// SIMATIC S7-200 SMART project (STEP 7-Micro/WIN SMART), CPU ST20

SYMBOL_TABLE 表格 1
Btn_set_Charge   V536.3
Calc_Temp_Real   VD700    // 计算中间暂存区 (DInt/Real)
Comm_State_Counter VB548    // 串口发送逻辑切换计数器
Comm_State_Counter1 VB549
HMI_IP_Apply     V536.2   // HMI 确认修改 IP 按钮
HMI_Start_Btn    V536.0   // HMI 手动开始按钮
HMI_Stop_Btn     V536.1   // HMI 手动停止按钮
Input_Current    VD504    // 实时输入电流 (A)
Input_Power      VD508    // 实时输入功率 (W)
Input_Voltage    VD500    // 实时输入电压 (V)
Output_Current   VD516    // 实时输出电流 (A)
Output_Voltage   VD512    // 实时输出电压 (V)
PLC_IP_Octet1    VB908    // PLC IP 地址第 1 段
PLC_IP_Octet2    VB909    // PLC IP 地址第 2 段
PLC_IP_Octet3    VB910    // PLC IP 地址第 3 段
PLC_IP_Octet4    VB911    // PLC IP 地址第 4 段
PN_In_Cmd        IB1160   // PN 接收自 1200: 远程启停指令
PN_In_SetI       ID1156   // PN 接收自 1200: 远程设定电流
PN_In_SetV       ID1152   // PN 接收自 1200: 远程设定电压
PN_Out_Curr      QD1156   // PN 发送给 1200: 输出电流
PN_Out_SetI      QD1164   // PN 发送给 1200: 当前设定电流
PN_Out_SetV      QD1160   // PN 发送给 1200: 当前设定电压
PN_Out_Status    QB1168   // PN 发送给 1200: 系统状态字节
PN_Out_Volt      QD1152   // PN 发送给 1200: 输出电压
Set_Current      VD532    // HMI 设定电流值 (默认 15.0)
Set_Voltage      VD528    // HMI 设定电压值 (默认 54.0)
Status_Bat_FB    V537.2   // 电池接入状态 (对应 Q0.1)
Status_Fault_FB  V537.1   // 系统故障状态 (对应 Q0.2)
Status_Run_FB    V537.0   // 充电运行状态 (对应 Q0.0)
Status_开关机标志     V537.3
Temp_T1          VD520    // 模块温度 T1 (℃)
Temp_T2          VD524    // 模块温度 T2 (℃)
发送数据             VB600    // 串口发送缓冲区起始 (长度 13)
启动接收并存入_VB550    VB550
END_SYMBOL_TABLE

SYMBOL_TABLE 系统符号
Always_On        SM0.0    // 始终接通
First_Scan_On    SM0.1    // 仅在第一个扫描周期时接通
P0_Config        SMB30    // 组态端口 0 通信：奇偶校验、每个字符的数据位数、波特率和协议
P0_Ctrl_Rcv      SMB87    // 接收消息控制
P0_End_Char      SMB89    // 消息结束字符
P0_Timeout       SMW92    // 字符间/消息定时器超时值，以毫秒为单位指定
P0_Max_Char      SMB94    // 要接收的最大字符数（1 到 255 字节）
END_SYMBOL_TABLE

ORGANIZATION_BLOCK MAIN:OB1
TITLE=
BEGIN
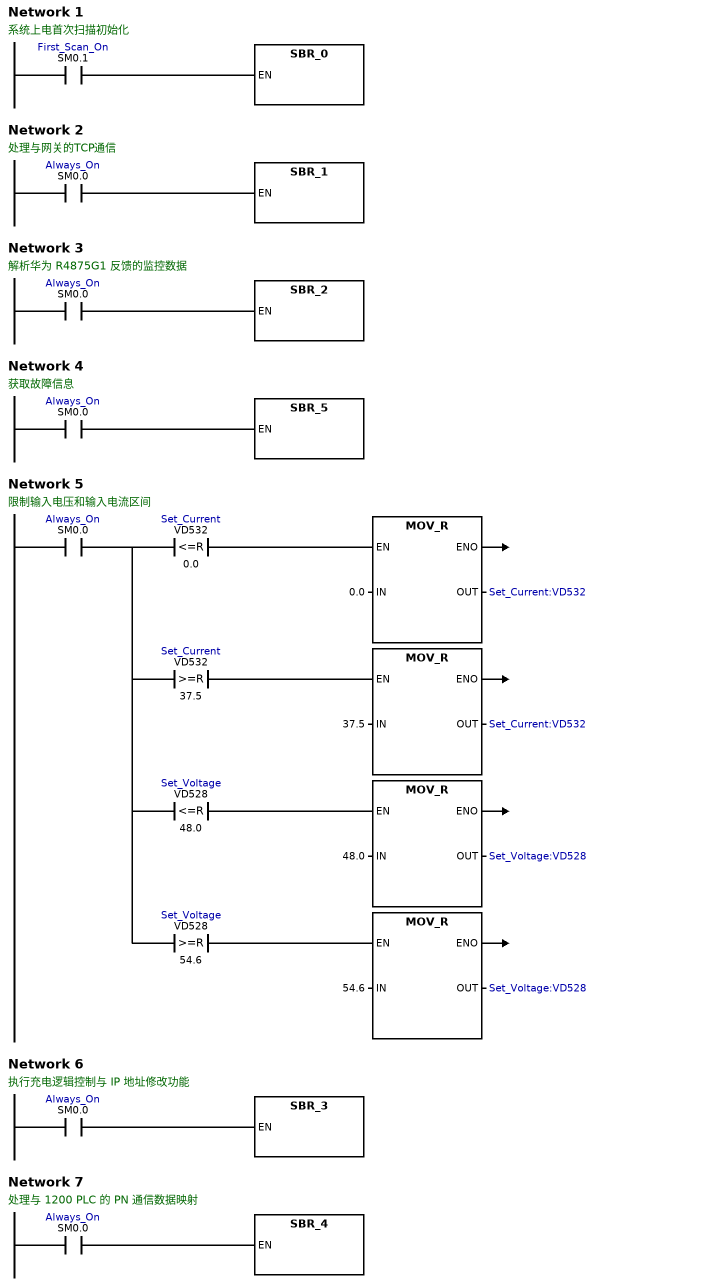
Network 1
//  系统上电首次扫描初始化
// 载入首次扫描标志位
// 调用初始化子程序
LD     First_Scan_On:SM0.1
CALL   SBR_0:SBR0
Network 2
//  处理与网关的TCP通信
// 始终接通
// 调用通信子程序
LD     Always_On:SM0.0
CALL   SBR_1:SBR1
Network 3
//  解析华为 R4875G1 反馈的监控数据
// 始终接通
// 调用解析子程序
LD     Always_On:SM0.0
CALL   SBR_2:SBR2
Network 4
// 获取故障信息
// 始终接通
// 调用获取故障程序
LD     Always_On:SM0.0
CALL   SBR_5:SBR5
Network 5
// 限制输入电压和输入电流区间
LD     Always_On:SM0.0
LPS
AR<=   Set_Current:VD532, 0.0
MOVR   0.0, Set_Current:VD532
LRD
AR>=   Set_Current:VD532, 37.5
MOVR   37.5, Set_Current:VD532
LRD
AR<=   Set_Voltage:VD528, 48.0
MOVR   48.0, Set_Voltage:VD528
LPP
AR>=   Set_Voltage:VD528, 54.6
MOVR   54.6, Set_Voltage:VD528
Network 6
//  执行充电逻辑控制与 IP 地址修改功能
// 始终接通
// 调用控制子程序
LD     Always_On:SM0.0
CALL   SBR_3:SBR3
Network 7
//  处理与 1200 PLC 的 PN 通信数据映射
// 始终接通
// 调用通信映射子程序
LD     Always_On:SM0.0
CALL   SBR_4:SBR4
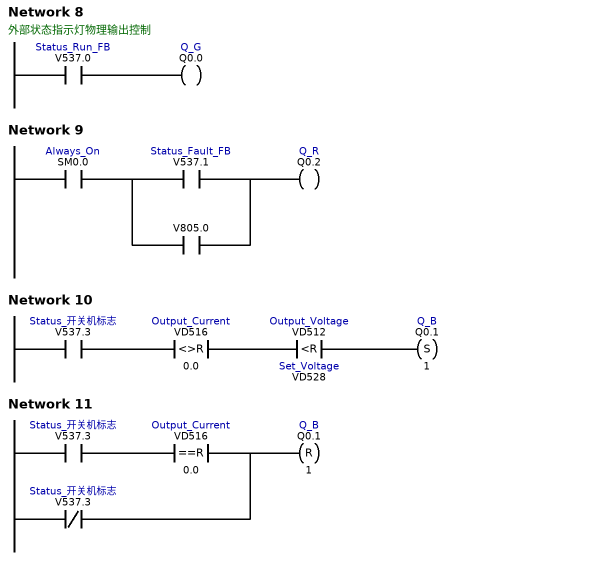
Network 8
//  外部状态指示灯物理输出控制
// 检查运行状态位
// 输出 Q0.0 绿灯: 充电运行
LD     Status_Run_FB:V537.0
=      Q_G:Q0.0
Network 9
// 检查故障状态位
// 输出 Q0.2 红灯: 系统故障
LD     Always_On:SM0.0
LD     Status_Fault_FB:V537.1
O      V805.0
ALD
=      Q_R:Q0.2
Network 10
// 检查电池接入位 (特殊标记：需用户自行完善)
// 输出 Q0.1 蓝灯: 电池接入
LD     Status_开关机标志:V537.3
AR<>   Output_Current:VD516, 0.0
AR<    Output_Voltage:VD512, Set_Voltage:VD528
S      Q_B:Q0.1, 1
Network 11
// 检查电池接入位 (特殊标记：需用户自行完善)
// 输出 Q0.1 蓝灯: 电池接入
LD     Status_开关机标志:V537.3
AR=    Output_Current:VD516, 0.0
ON     Status_开关机标志:V537.3
R      Q_B:Q0.1, 1
END_ORGANIZATION_BLOCK

SUBROUTINE_BLOCK SBR_0:SBR0
TITLE=初始化子程序
BEGIN
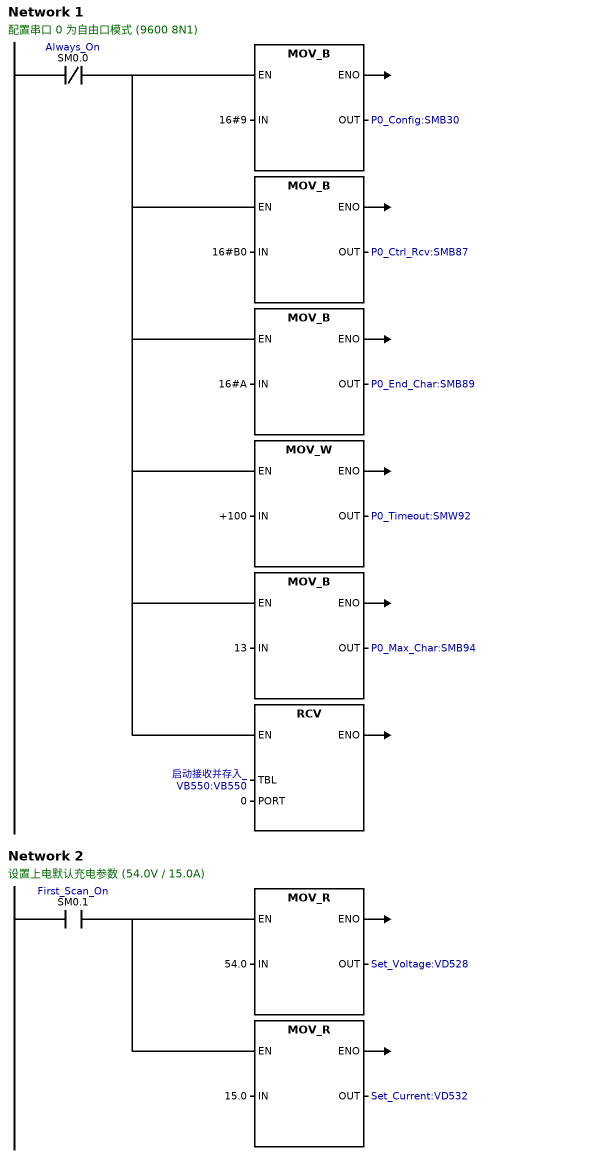
Network 1
//  配置串口 0 为自由口模式 (9600 8N1)
// 始终接通
// 端口 0: 9600, 8, N, 1, 自由口
// 设置接收控制: 允许接收, 超时结束
// 设置结束符 (0x0A)
// 设置接收超时 100ms
// 设置最大接收长度 13 字节
// 启动接收并存入 VB550
LDN    Always_On:SM0.0
MOVB   16#9, P0_Config:SMB30
MOVB   16#B0, P0_Ctrl_Rcv:SMB87
MOVB   16#A, P0_End_Char:SMB89
MOVW   +100, P0_Timeout:SMW92
MOVB   13, P0_Max_Char:SMB94
RCV    启动接收并存入_VB550:VB550, 0
Network 2
//  设置上电默认充电参数 (54.0V / 15.0A)
// 首次扫描
// 默认设定电压 54.0V
// 默认设定电流 15.0A
LD     First_Scan_On:SM0.1
MOVR   54.0, Set_Voltage:VD528
MOVR   15.0, Set_Current:VD532
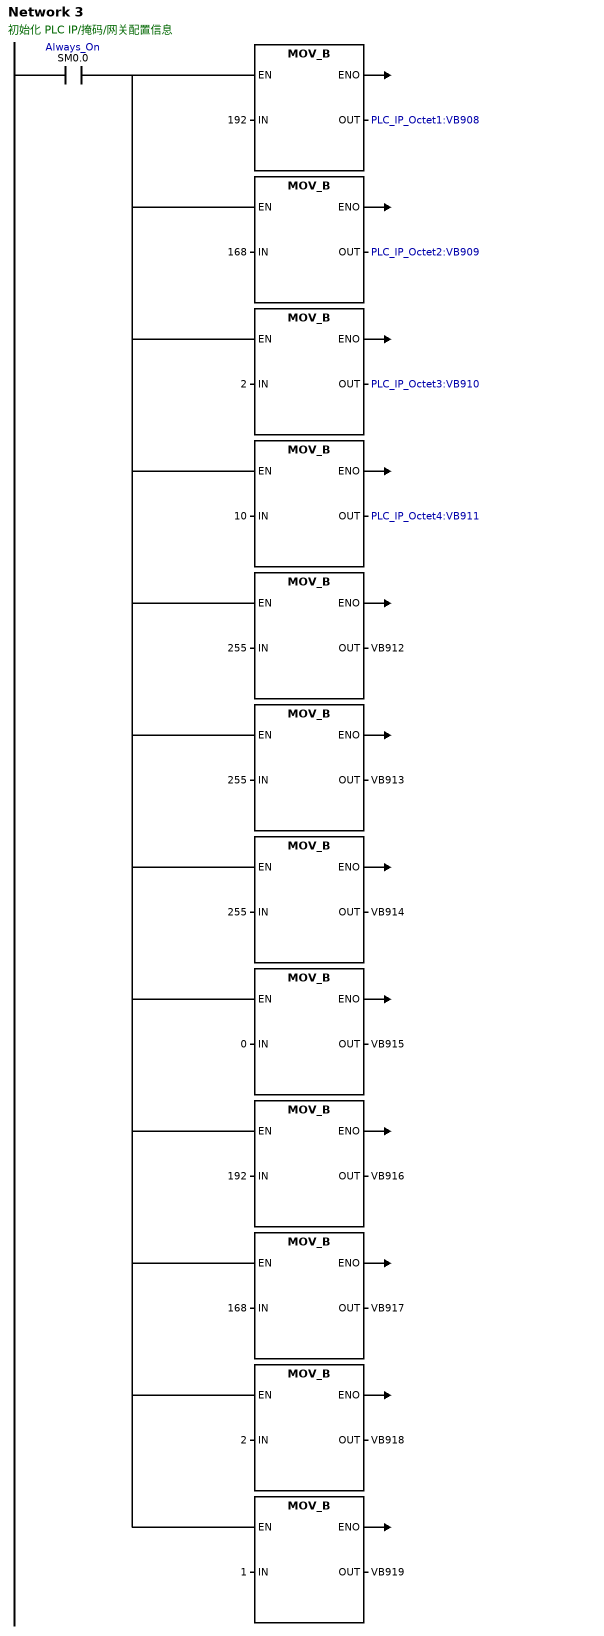
Network 3
//  初始化 PLC IP/掩码/网关配置信息
// 首次扫描
// IP 第一段
// IP 第二段
// IP 第三段
// IP 第四段
// 掩码第一段
// 掩码第二段
// 掩码第三段
// 掩码第四段
// 网关第一段
// 网关第二段
// 网关第三段
// 网关第四段
LD     Always_On:SM0.0
MOVB   192, PLC_IP_Octet1:VB908
MOVB   168, PLC_IP_Octet2:VB909
MOVB   2, PLC_IP_Octet3:VB910
MOVB   10, PLC_IP_Octet4:VB911
MOVB   255, VB912
MOVB   255, VB913
MOVB   255, VB914
MOVB   0, VB915
MOVB   192, VB916
MOVB   168, VB917
MOVB   2, VB918
MOVB   1, VB919
END_SUBROUTINE_BLOCK

SUBROUTINE_BLOCK SBR_1:SBR1
TITLE=TCP通信 - 华为协议
BEGIN
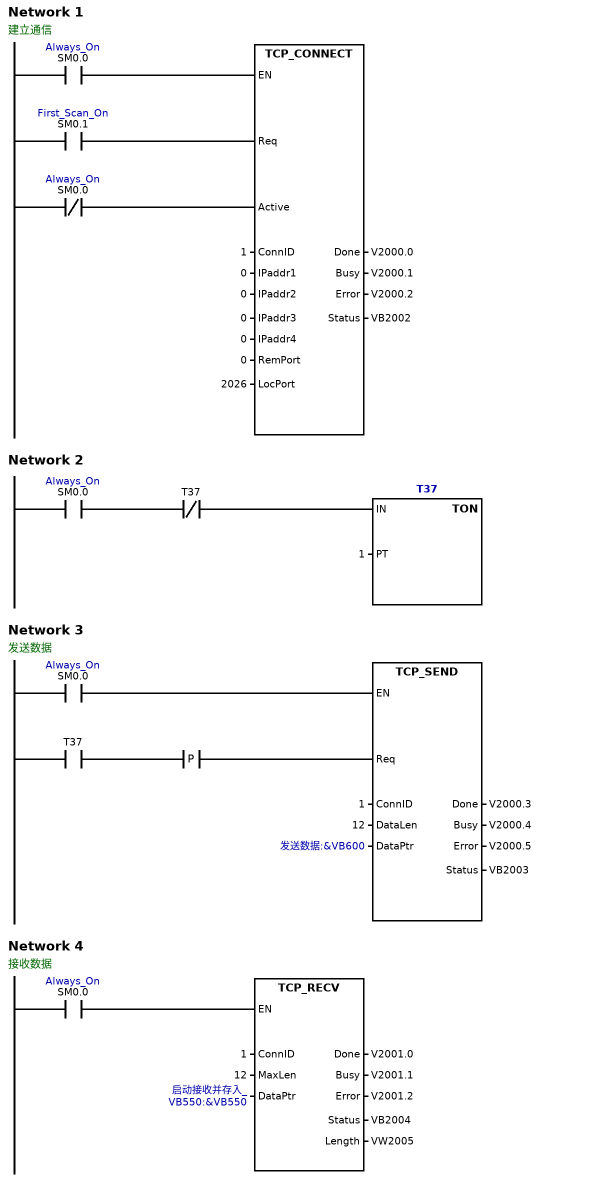
Network 1
// 建立通信
LD     Always_On:SM0.0
=      L60.0
LD     First_Scan_On:SM0.1
=      L63.7
LDN    Always_On:SM0.0
=      L63.6
LD     L60.0
CALL   TCP_CONNECT:SBR6, L63.7, L63.6, 1, 0, 0, 0, 0, 0, 2026, V2000.0, V2000.1, V2000.2, VB2002
Network 2
LD     Always_On:SM0.0
AN     T37
TON    T37, 1
Network 3
// 发送数据
LD     Always_On:SM0.0
=      L60.0
LD     T37
EU
=      L63.7
LD     L60.0
CALL   TCP_SEND:SBR7, L63.7, 1, 12, &发送数据:VB600, V2000.3, V2000.4, V2000.5, VB2003
Network 4
// 接收数据
LD     Always_On:SM0.0
CALL   TCP_RECV:SBR8, 1, 12, &启动接收并存入_VB550:VB550, V2001.0, V2001.1, V2001.2, VB2004, VW2005
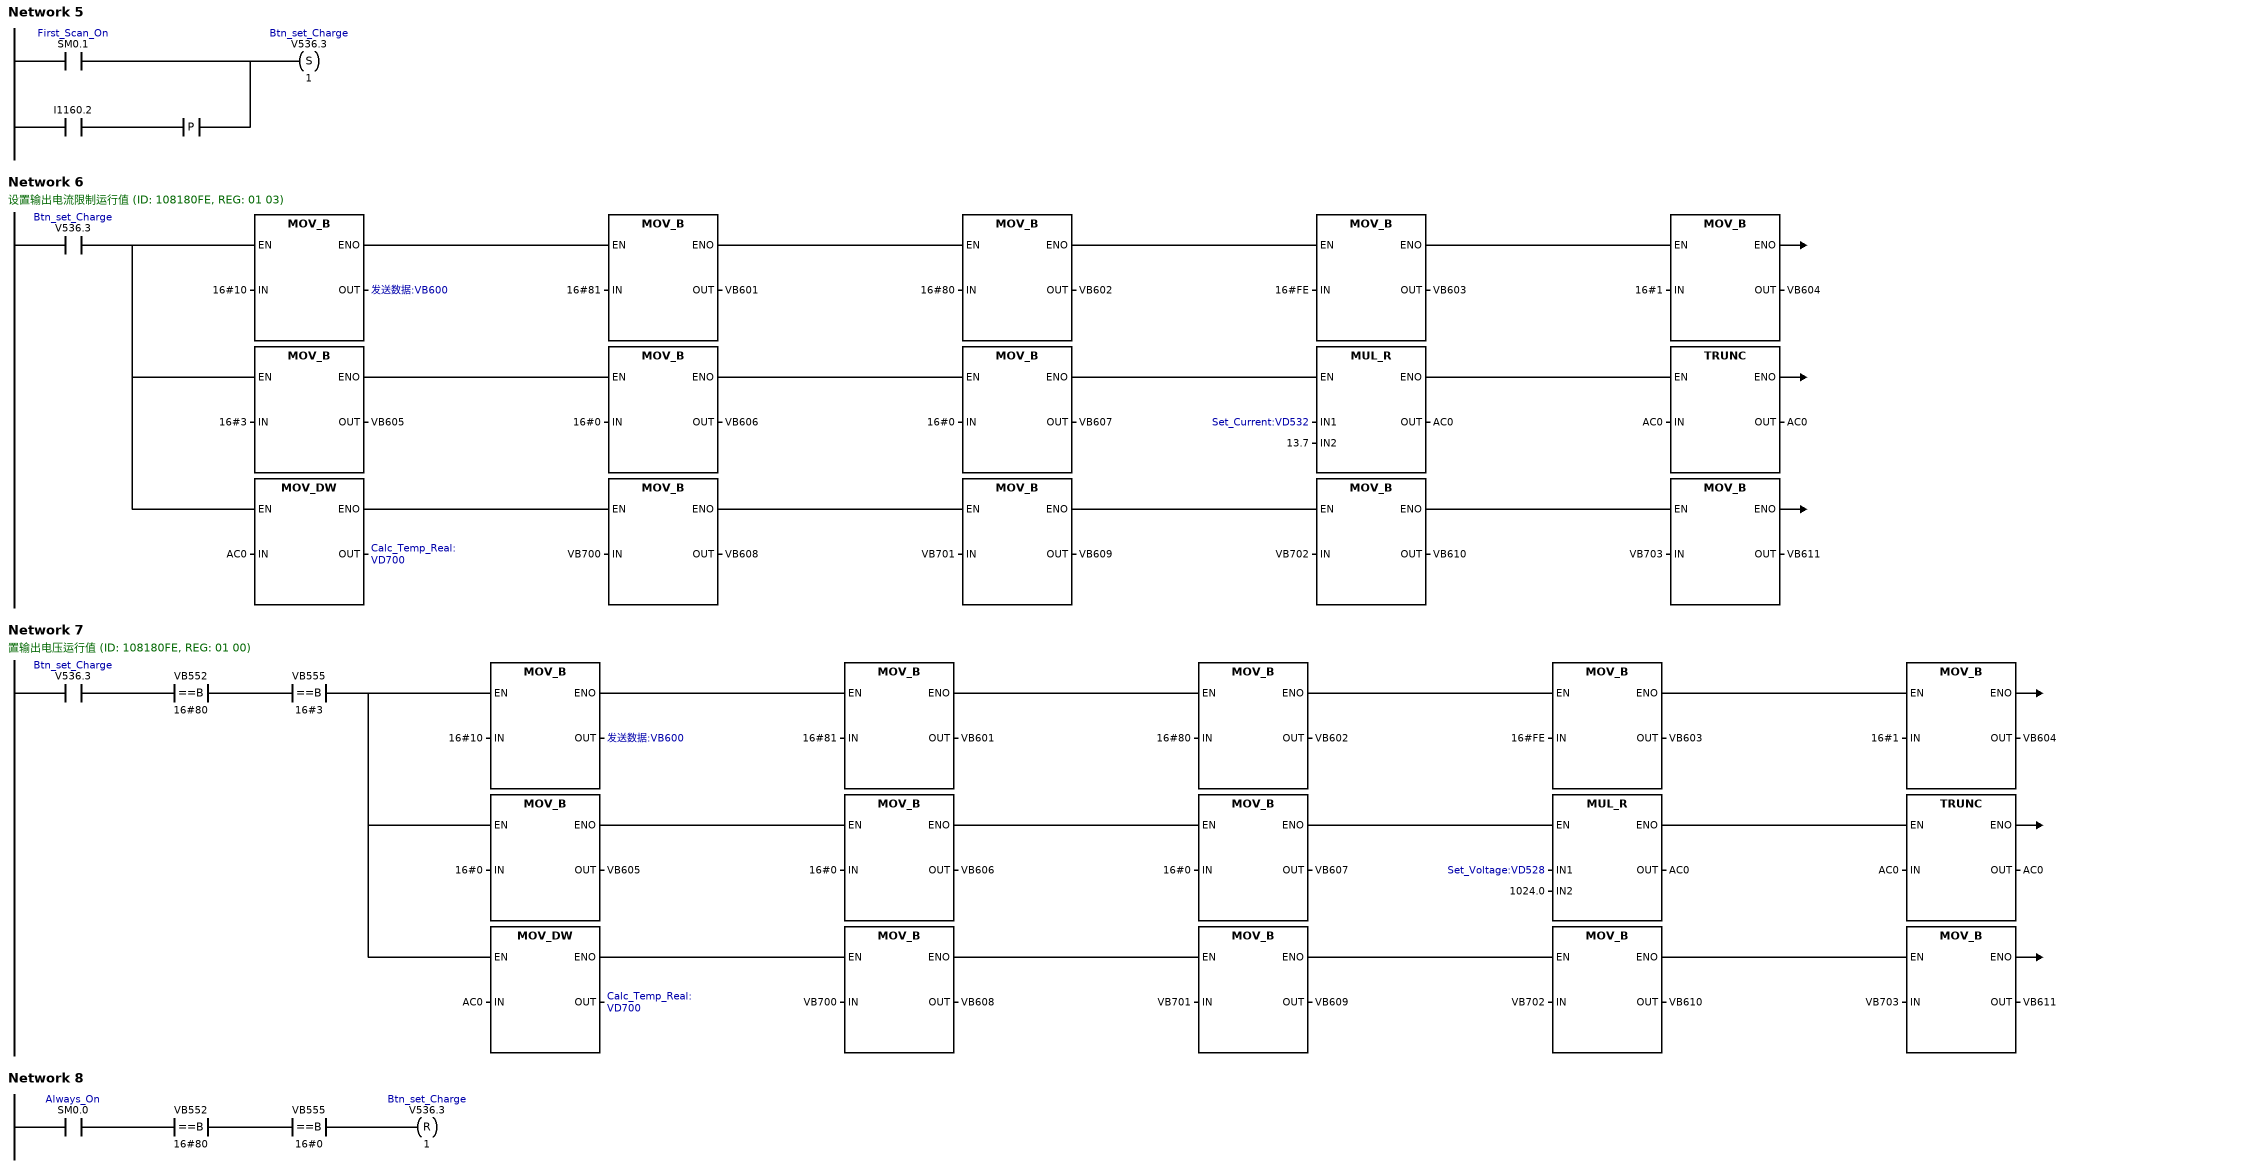
Network 5
LD     First_Scan_On:SM0.1
LD     I1160.2
EU
OLD
S      Btn_set_Charge:V536.3, 1
Network 6
//  设置输出电流限制运行值 (ID: 108180FE, REG: 01 03)
LD     Btn_set_Charge:V536.3
LPS
MOVB   16#10, 发送数据:VB600
AENO
MOVB   16#81, VB601
AENO
MOVB   16#80, VB602
AENO
MOVB   16#FE, VB603
AENO
MOVB   16#1, VB604
LRD
MOVB   16#3, VB605
AENO
MOVB   16#0, VB606
AENO
MOVB   16#0, VB607
AENO
MOVR   Set_Current:VD532, AC0
AENO
*R     13.7, AC0
AENO
TRUNC  AC0, AC0
LPP
MOVD   AC0, Calc_Temp_Real:VD700
AENO
MOVB   VB700, VB608
AENO
MOVB   VB701, VB609
AENO
MOVB   VB702, VB610
AENO
MOVB   VB703, VB611
Network 7
// 置输出电压运行值 (ID: 108180FE, REG: 01 00)
// 状态 3：处理启停
// 若状态计数器等于 1
// CAN ID Byte 3
// CAN ID Byte 2
// CAN ID Byte 1
// CAN ID Byte 0 (修正为 FE)
// 华为数据 Byte 0
// 华为数据 Byte 1 (寄存器 01 00)
// 华为数据 Byte 2
// 华为数据 Byte 3
// 载入 HMI 设定电压值
// 乘以 1024
// 转换为双整数
// 暂存至 VD700
// 填充设定值字节 4 (大端)
// 填充设定值字节 5
// 填充设定值字节 6
// 填充设定值字节 7
LD     Btn_set_Charge:V536.3
AB=    VB552, 16#80
AB=    VB555, 16#3
LPS
MOVB   16#10, 发送数据:VB600
AENO
MOVB   16#81, VB601
AENO
MOVB   16#80, VB602
AENO
MOVB   16#FE, VB603
AENO
MOVB   16#1, VB604
LRD
MOVB   16#0, VB605
AENO
MOVB   16#0, VB606
AENO
MOVB   16#0, VB607
AENO
MOVR   Set_Voltage:VD528, AC0
AENO
*R     1024.0, AC0
AENO
TRUNC  AC0, AC0
LPP
MOVD   AC0, Calc_Temp_Real:VD700
AENO
MOVB   VB700, VB608
AENO
MOVB   VB701, VB609
AENO
MOVB   VB702, VB610
AENO
MOVB   VB703, VB611
Network 8
LD     Always_On:SM0.0
AB=    VB552, 16#80
AB=    VB555, 16#0
R      Btn_set_Charge:V536.3, 1
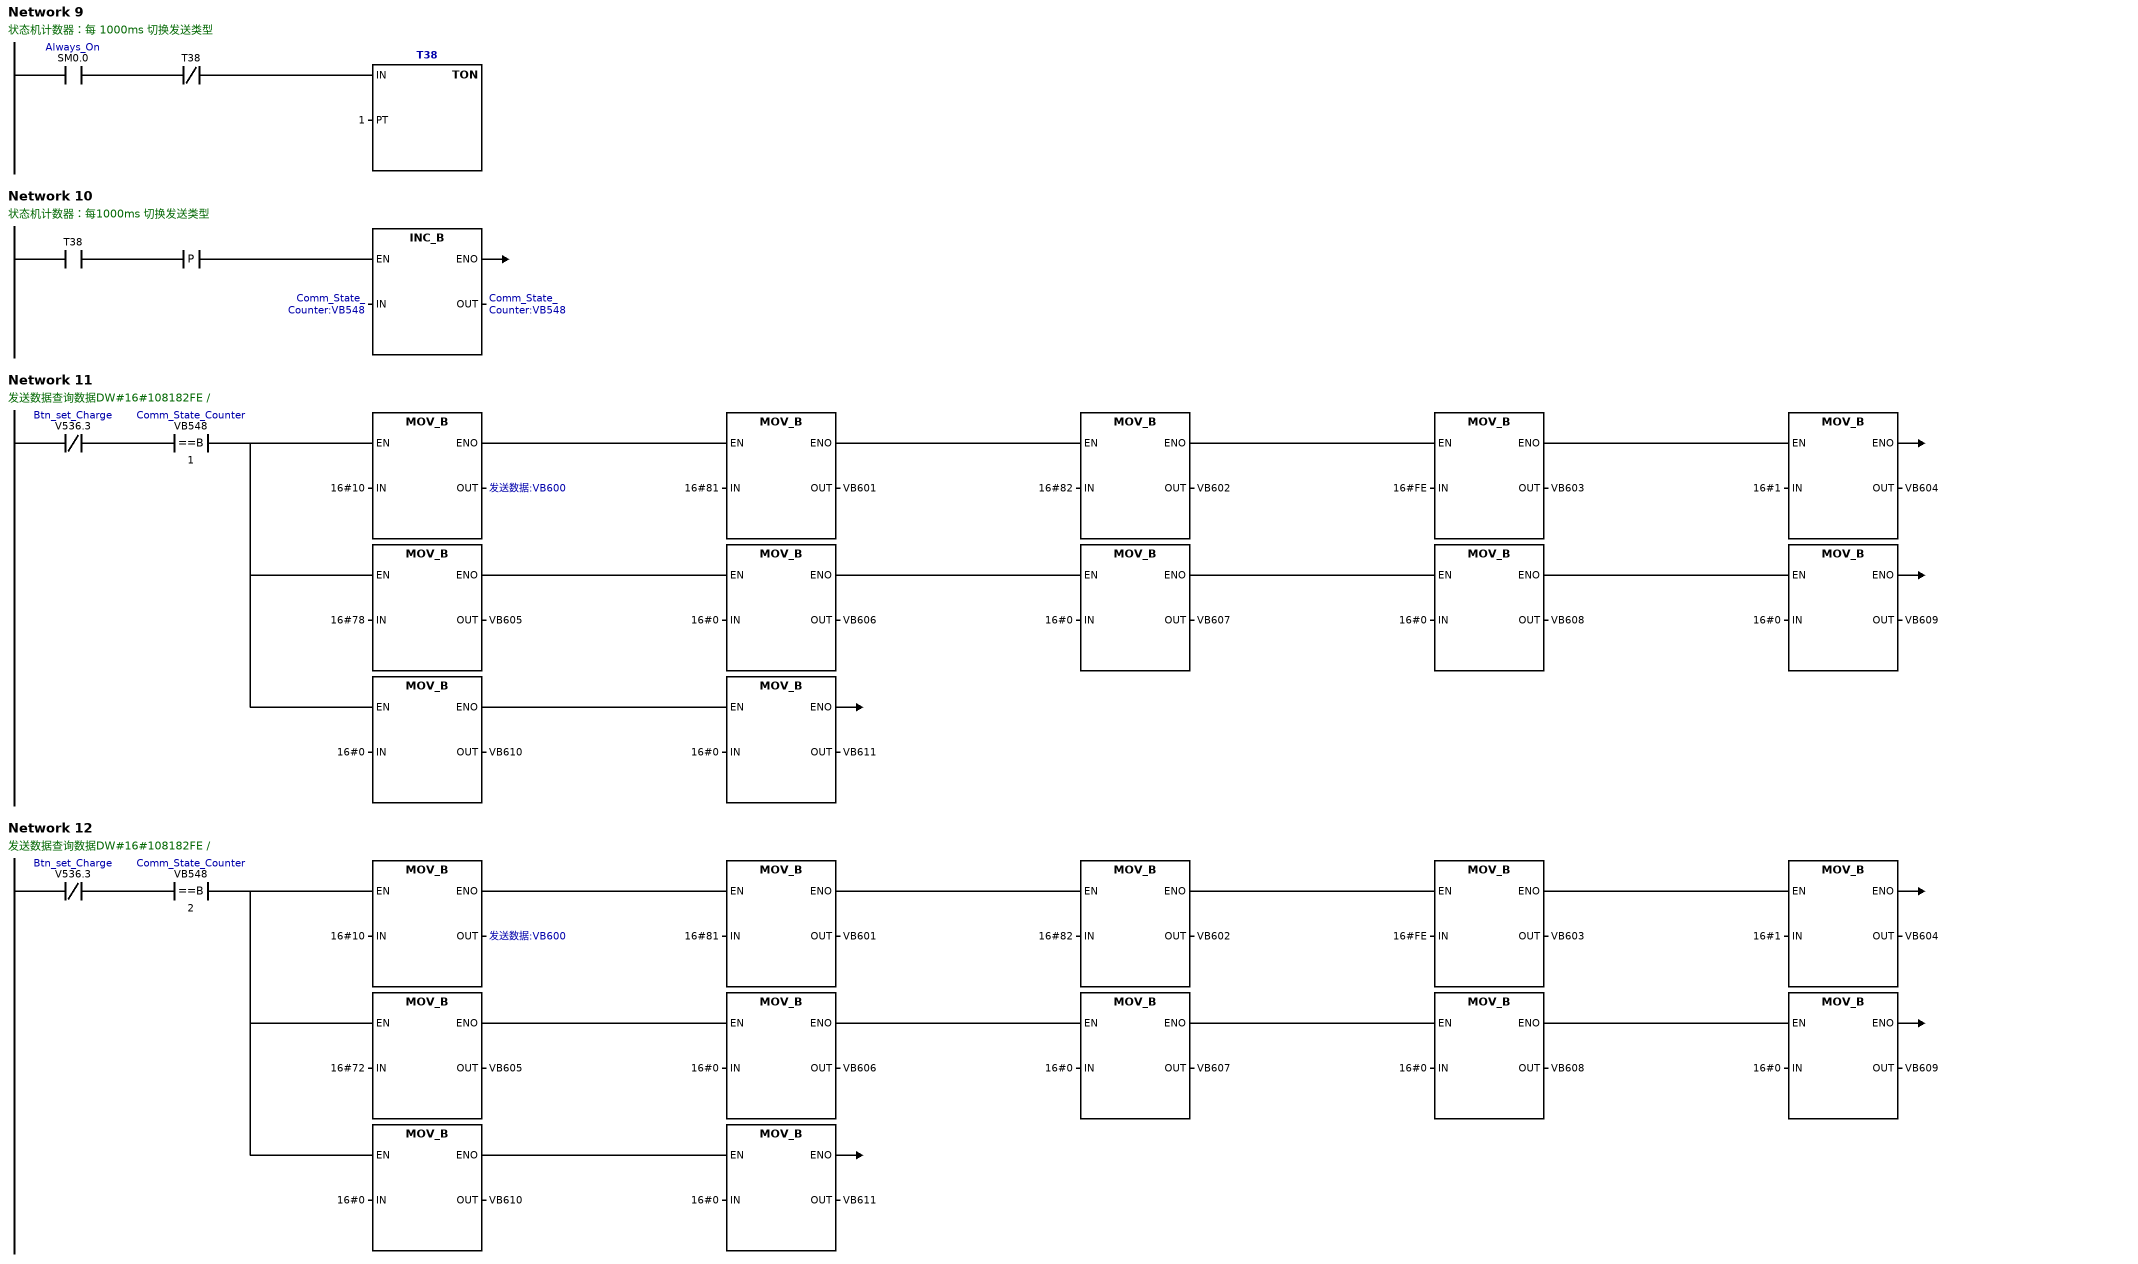
Network 9
// 状态机计数器：每 1000ms 切换发送类型
LD     Always_On:SM0.0
AN     T38
TON    T38, 1
Network 10
//  状态机计数器：每1000ms 切换发送类型
// 1s 脉冲
// 上升沿
// VB548 状态计数器自增
LD     T38
EU
INCB   Comm_State_Counter:VB548
Network 11
// 发送数据查询数据DW#16#108182FE
// 
// 状态 3：处理启停
// 若状态计数器等于 1 
// ID 3
// ID 2
// ID 1
// ID 0 (FE)
// Byte 0
// Byte 1 
// Byte 2
// Byte 3
// Byte 4
// Byte 5
// Byte 6
// Byte 7
LDN    Btn_set_Charge:V536.3
AB=    Comm_State_Counter:VB548, 1
LPS
MOVB   16#10, 发送数据:VB600
AENO
MOVB   16#81, VB601
AENO
MOVB   16#82, VB602
AENO
MOVB   16#FE, VB603
AENO
MOVB   16#1, VB604
LRD
MOVB   16#78, VB605
AENO
MOVB   16#0, VB606
AENO
MOVB   16#0, VB607
AENO
MOVB   16#0, VB608
AENO
MOVB   16#0, VB609
LPP
MOVB   16#0, VB610
AENO
MOVB   16#0, VB611
Network 12
// 发送数据查询数据DW#16#108182FE
// 
// 状态 3：处理启停
// 若状态计数器等于 2 
// ID 3
// ID 2
// ID 1
// ID 0 (FE)
// Byte 0
// Byte 1 
// Byte 2
// Byte 3
// Byte 4
// Byte 5
// Byte 6
// Byte 7
LDN    Btn_set_Charge:V536.3
AB=    Comm_State_Counter:VB548, 2
LPS
MOVB   16#10, 发送数据:VB600
AENO
MOVB   16#81, VB601
AENO
MOVB   16#82, VB602
AENO
MOVB   16#FE, VB603
AENO
MOVB   16#1, VB604
LRD
MOVB   16#72, VB605
AENO
MOVB   16#0, VB606
AENO
MOVB   16#0, VB607
AENO
MOVB   16#0, VB608
AENO
MOVB   16#0, VB609
LPP
MOVB   16#0, VB610
AENO
MOVB   16#0, VB611
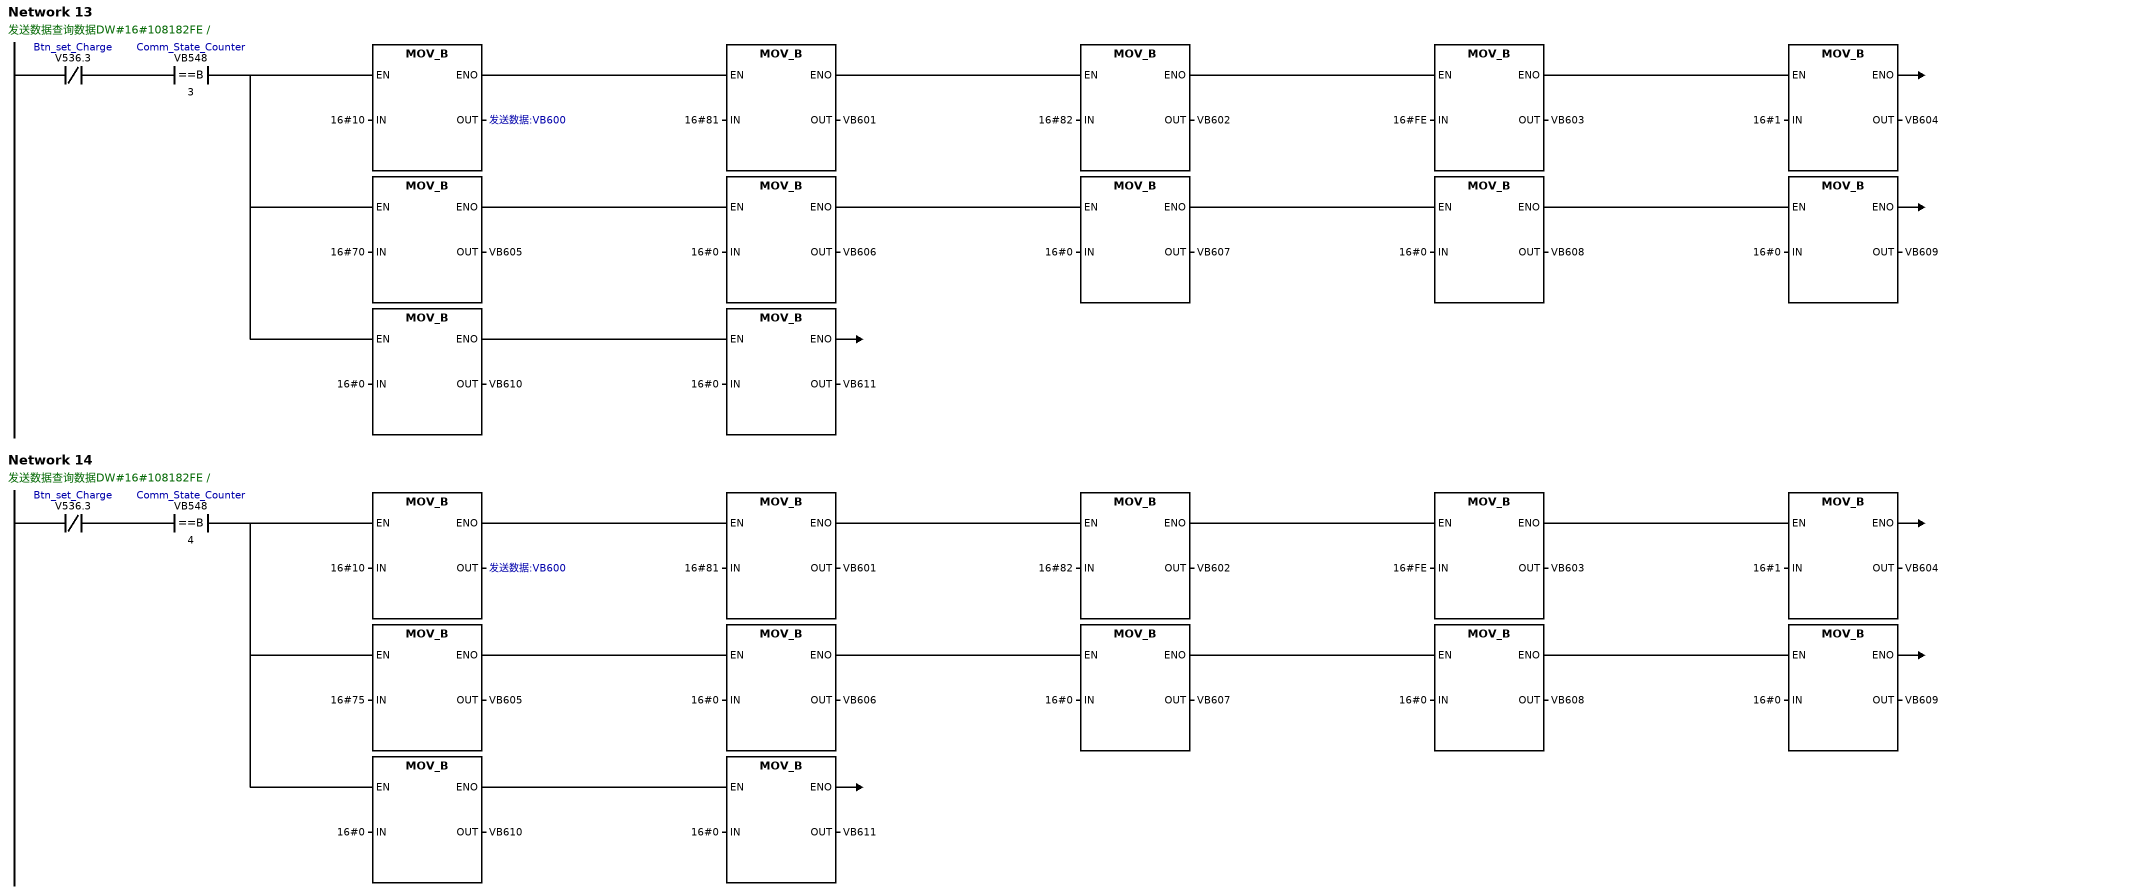
Network 13
// 发送数据查询数据DW#16#108182FE
// 
// 状态 3：处理启停
// 若状态计数器等于 3 
// ID 3
// ID 2
// ID 1
// ID 0 (FE)
// Byte 0
// Byte 1 
// Byte 2
// Byte 3
// Byte 4
// Byte 5
// Byte 6
// Byte 7
LDN    Btn_set_Charge:V536.3
AB=    Comm_State_Counter:VB548, 3
LPS
MOVB   16#10, 发送数据:VB600
AENO
MOVB   16#81, VB601
AENO
MOVB   16#82, VB602
AENO
MOVB   16#FE, VB603
AENO
MOVB   16#1, VB604
LRD
MOVB   16#70, VB605
AENO
MOVB   16#0, VB606
AENO
MOVB   16#0, VB607
AENO
MOVB   16#0, VB608
AENO
MOVB   16#0, VB609
LPP
MOVB   16#0, VB610
AENO
MOVB   16#0, VB611
Network 14
// 发送数据查询数据DW#16#108182FE
// 
// 状态 3：处理启停
// 若状态计数器等于 4
// ID 2
// ID 1
// ID 0 (FE)
// Byte 0
// Byte 1 
// Byte 2
// Byte 3
// Byte 4
// Byte 5
// Byte 6
// Byte 7
LDN    Btn_set_Charge:V536.3
AB=    Comm_State_Counter:VB548, 4
LPS
MOVB   16#10, 发送数据:VB600
AENO
MOVB   16#81, VB601
AENO
MOVB   16#82, VB602
AENO
MOVB   16#FE, VB603
AENO
MOVB   16#1, VB604
LRD
MOVB   16#75, VB605
AENO
MOVB   16#0, VB606
AENO
MOVB   16#0, VB607
AENO
MOVB   16#0, VB608
AENO
MOVB   16#0, VB609
LPP
MOVB   16#0, VB610
AENO
MOVB   16#0, VB611
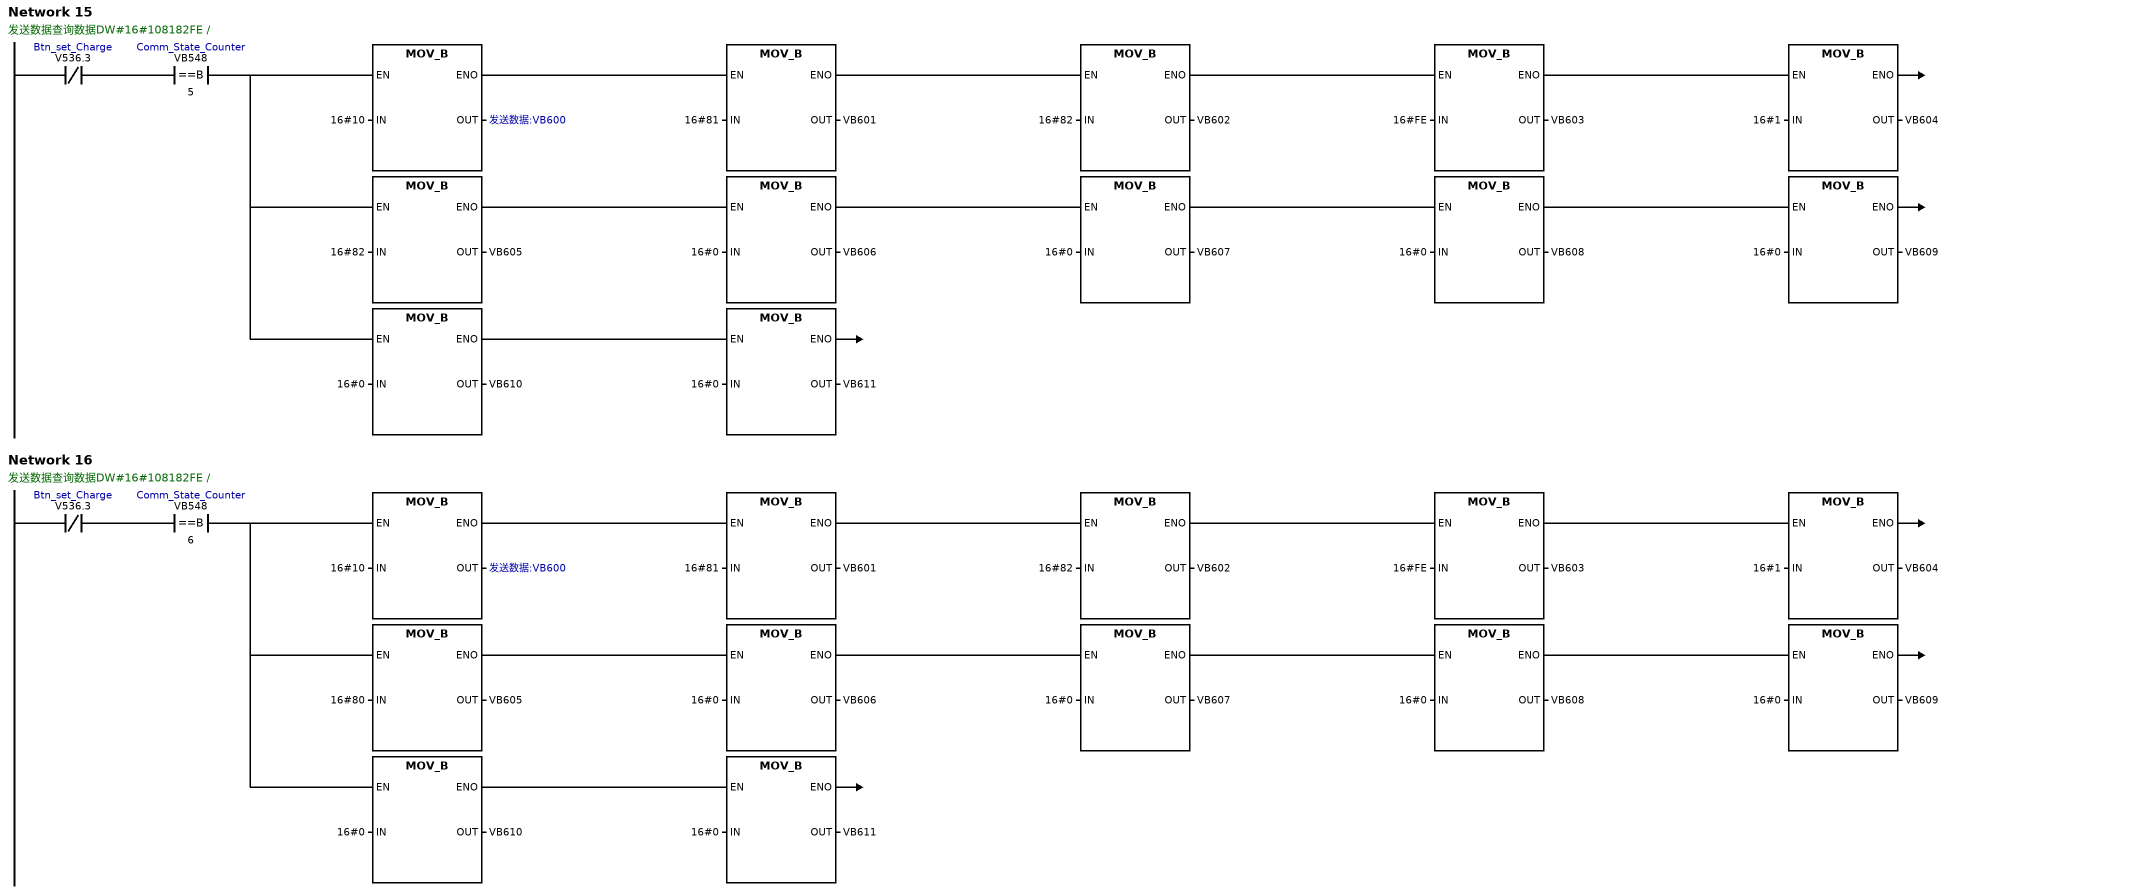
Network 15
// 发送数据查询数据DW#16#108182FE
// 
// 状态 3：处理启停
// 若状态计数器等于 5
// ID 2
// ID 1
// ID 0 (FE)
// Byte 0
// Byte 1 
// Byte 2
// Byte 3
// Byte 4
// Byte 5
// Byte 6
// Byte 7
LDN    Btn_set_Charge:V536.3
AB=    Comm_State_Counter:VB548, 5
LPS
MOVB   16#10, 发送数据:VB600
AENO
MOVB   16#81, VB601
AENO
MOVB   16#82, VB602
AENO
MOVB   16#FE, VB603
AENO
MOVB   16#1, VB604
LRD
MOVB   16#82, VB605
AENO
MOVB   16#0, VB606
AENO
MOVB   16#0, VB607
AENO
MOVB   16#0, VB608
AENO
MOVB   16#0, VB609
LPP
MOVB   16#0, VB610
AENO
MOVB   16#0, VB611
Network 16
// 发送数据查询数据DW#16#108182FE
// 
// 状态 3：处理启停
// 若状态计数器等于 6
// ID 2
// ID 1
// ID 0 (FE)
// Byte 0
// Byte 1 
// Byte 2
// Byte 3
// Byte 4
// Byte 5
// Byte 6
// Byte 7
LDN    Btn_set_Charge:V536.3
AB=    Comm_State_Counter:VB548, 6
LPS
MOVB   16#10, 发送数据:VB600
AENO
MOVB   16#81, VB601
AENO
MOVB   16#82, VB602
AENO
MOVB   16#FE, VB603
AENO
MOVB   16#1, VB604
LRD
MOVB   16#80, VB605
AENO
MOVB   16#0, VB606
AENO
MOVB   16#0, VB607
AENO
MOVB   16#0, VB608
AENO
MOVB   16#0, VB609
LPP
MOVB   16#0, VB610
AENO
MOVB   16#0, VB611
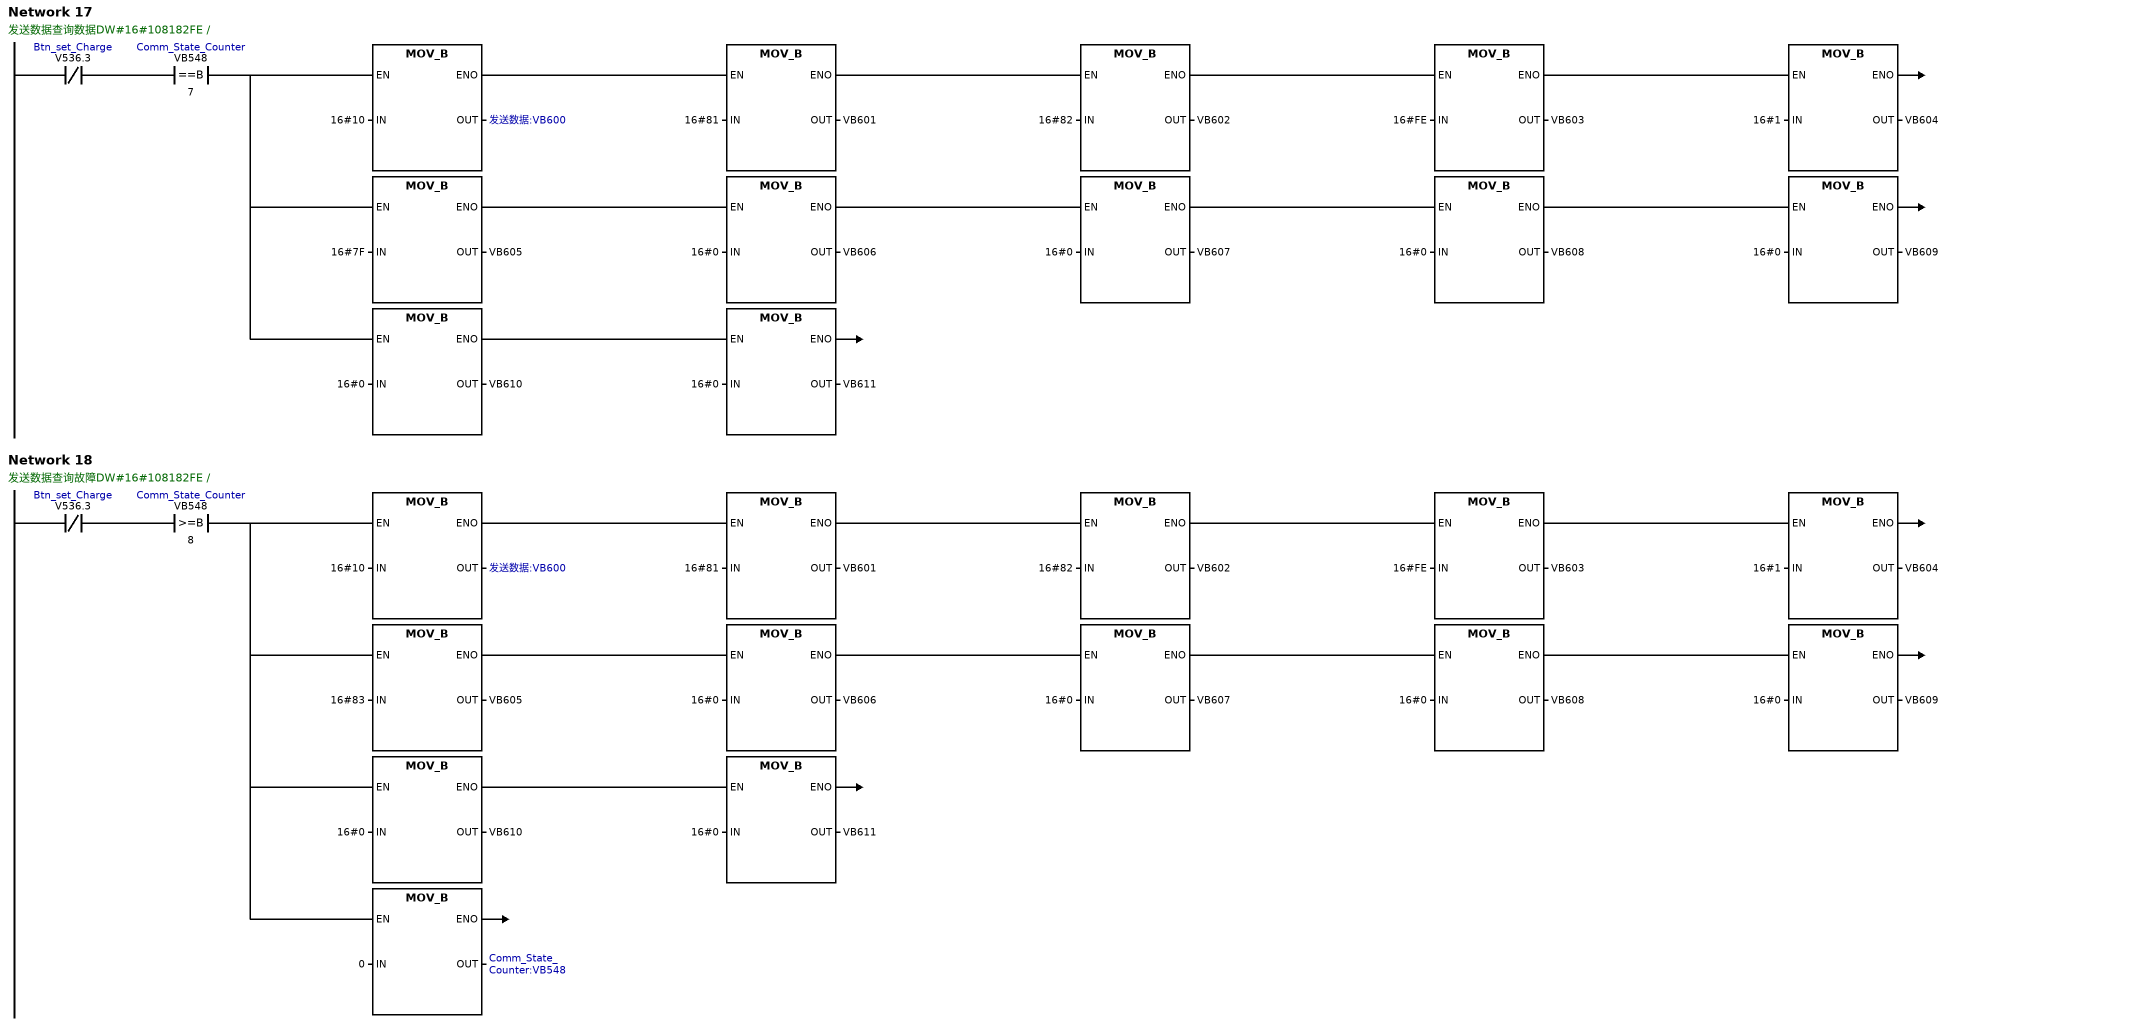
Network 17
// 发送数据查询数据DW#16#108182FE
// 
// 状态 3：处理启停
// 若状态计数器等于 7
// ID 2
// ID 1
// ID 0 (FE)
// Byte 0
// Byte 1 
// Byte 2
// Byte 3
// Byte 4
// Byte 5
// Byte 6
// Byte 7
LDN    Btn_set_Charge:V536.3
AB=    Comm_State_Counter:VB548, 7
LPS
MOVB   16#10, 发送数据:VB600
AENO
MOVB   16#81, VB601
AENO
MOVB   16#82, VB602
AENO
MOVB   16#FE, VB603
AENO
MOVB   16#1, VB604
LRD
MOVB   16#7F, VB605
AENO
MOVB   16#0, VB606
AENO
MOVB   16#0, VB607
AENO
MOVB   16#0, VB608
AENO
MOVB   16#0, VB609
LPP
MOVB   16#0, VB610
AENO
MOVB   16#0, VB611
Network 18
// 发送数据查询故障DW#16#108182FE
// 
// 状态 3：处理启停
// 若状态计数器等于 8 
// 重置轮询计数器
// ID 3
// ID 2
// ID 1
// ID 0 (FE)
// Byte 0
// Byte 1 (寄存器 01 83)
// Byte 2
// Byte 3
// Byte 4
// Byte 5
// Byte 6
// Byte 7
LDN    Btn_set_Charge:V536.3
AB>=   Comm_State_Counter:VB548, 8
LPS
MOVB   16#10, 发送数据:VB600
AENO
MOVB   16#81, VB601
AENO
MOVB   16#82, VB602
AENO
MOVB   16#FE, VB603
AENO
MOVB   16#1, VB604
LRD
MOVB   16#83, VB605
AENO
MOVB   16#0, VB606
AENO
MOVB   16#0, VB607
AENO
MOVB   16#0, VB608
AENO
MOVB   16#0, VB609
LRD
MOVB   16#0, VB610
AENO
MOVB   16#0, VB611
LPP
MOVB   0, Comm_State_Counter:VB548
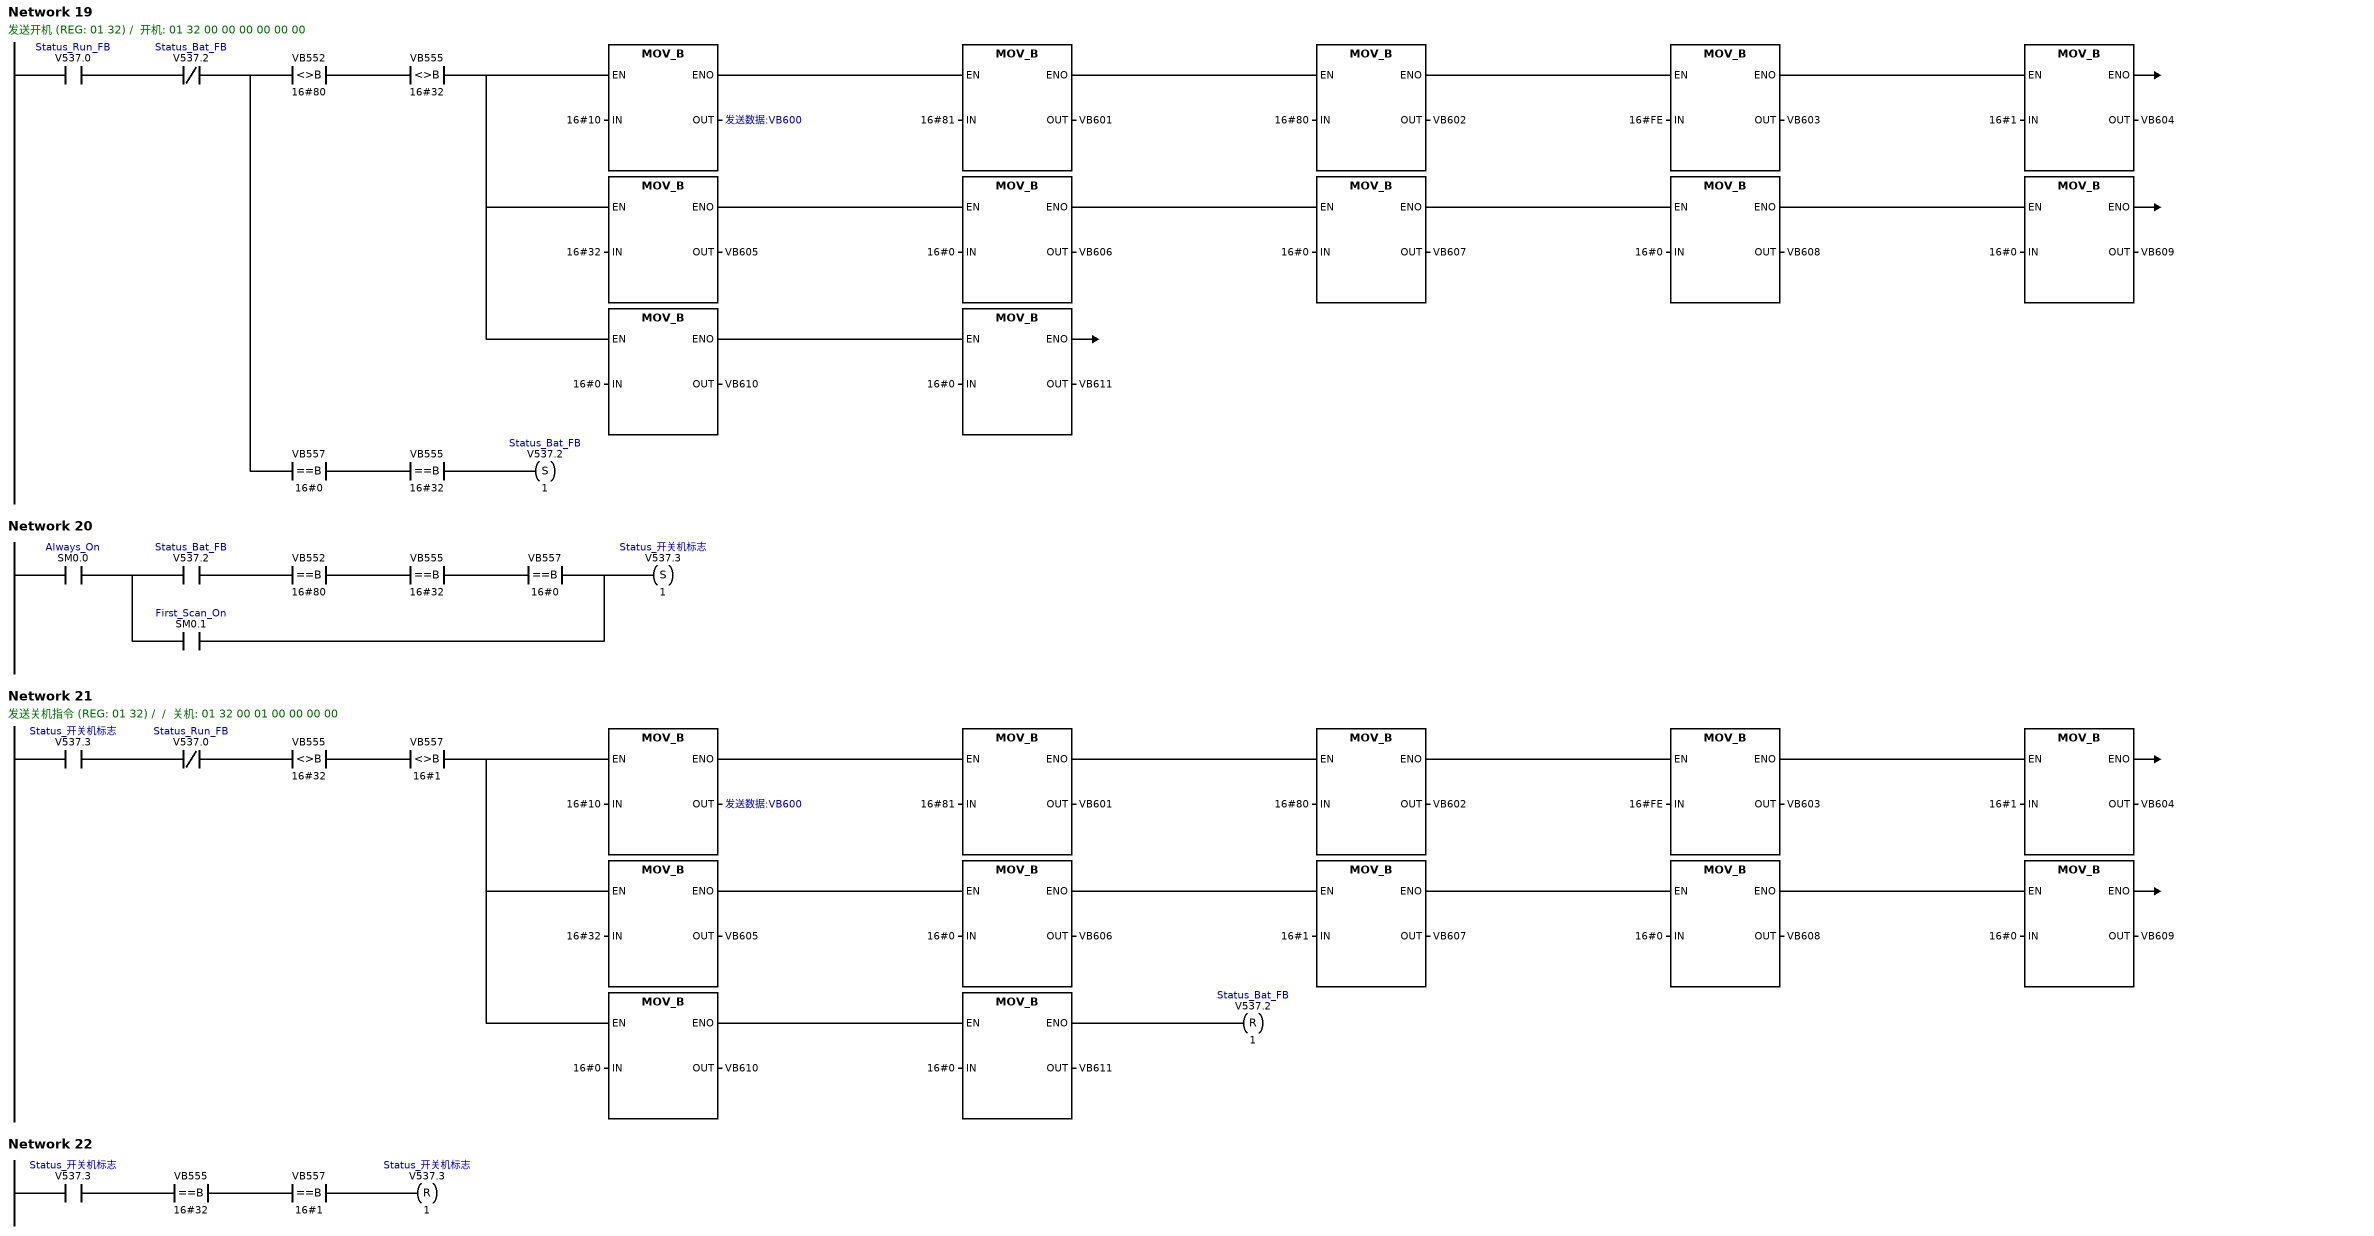
Network 19
// 发送开机 (REG: 01 32)
//  开机: 01 32 00 00 00 00 00 00
// 状态 3：处理启停
// 检查 ID 字节 1
// 参数 ID 为 0x32
// 参数 ID 为 0x00
// ID 3
// ID 2
// ID 1
// ID 0 (FE)
// Byte 0
// Byte 1 (寄存器 01 32)
// Byte 2
// 若运行标志为 0 (开机)
// Byte 4
// Byte 5
// Byte 6
// Byte 7
LD     Status_Run_FB:V537.0
AN     Status_Bat_FB:V537.2
LPS
AB<>   VB552, 16#80
AB<>   VB555, 16#32
LPS
MOVB   16#10, 发送数据:VB600
AENO
MOVB   16#81, VB601
AENO
MOVB   16#80, VB602
AENO
MOVB   16#FE, VB603
AENO
MOVB   16#1, VB604
LRD
MOVB   16#32, VB605
AENO
MOVB   16#0, VB606
AENO
MOVB   16#0, VB607
AENO
MOVB   16#0, VB608
AENO
MOVB   16#0, VB609
LPP
MOVB   16#0, VB610
AENO
MOVB   16#0, VB611
LPP
AB=    VB557, 16#0
AB=    VB555, 16#32
S      Status_Bat_FB:V537.2, 1
Network 20
LD     Always_On:SM0.0
LD     Status_Bat_FB:V537.2
AB=    VB552, 16#80
AB=    VB555, 16#32
AB=    VB557, 16#0
O      First_Scan_On:SM0.1
ALD
S      Status_开关机标志:V537.3, 1
Network 21
// 发送关机指令 (REG: 01 32)
// 
//  关机: 01 32 00 01 00 00 00 00
// 状态 3：处理启停
// 检查 ID 字节 1
// 参数 ID 为 0x32
// 参数 ID 为 0x01
// ID 3
// ID 2
// ID 1
// ID 0 (FE)
// Byte 0
// Byte 1 (寄存器 01 32)
// Byte 2
// 若运行标志为 1 (关机)
// Byte 4
// Byte 5
// Byte 6
// Byte 7
LD     Status_开关机标志:V537.3
AN     Status_Run_FB:V537.0
AB<>   VB555, 16#32
AB<>   VB557, 16#1
LPS
MOVB   16#10, 发送数据:VB600
AENO
MOVB   16#81, VB601
AENO
MOVB   16#80, VB602
AENO
MOVB   16#FE, VB603
AENO
MOVB   16#1, VB604
LRD
MOVB   16#32, VB605
AENO
MOVB   16#0, VB606
AENO
MOVB   16#1, VB607
AENO
MOVB   16#0, VB608
AENO
MOVB   16#0, VB609
LPP
MOVB   16#0, VB610
AENO
MOVB   16#0, VB611
AENO
R      Status_Bat_FB:V537.2, 1
Network 22
LD     Status_开关机标志:V537.3
AB=    VB555, 16#32
AB=    VB557, 16#1
R      Status_开关机标志:V537.3, 1
END_SUBROUTINE_BLOCK

SUBROUTINE_BLOCK SBR_2:SBR2
TITLE=数据解析子程序
BEGIN
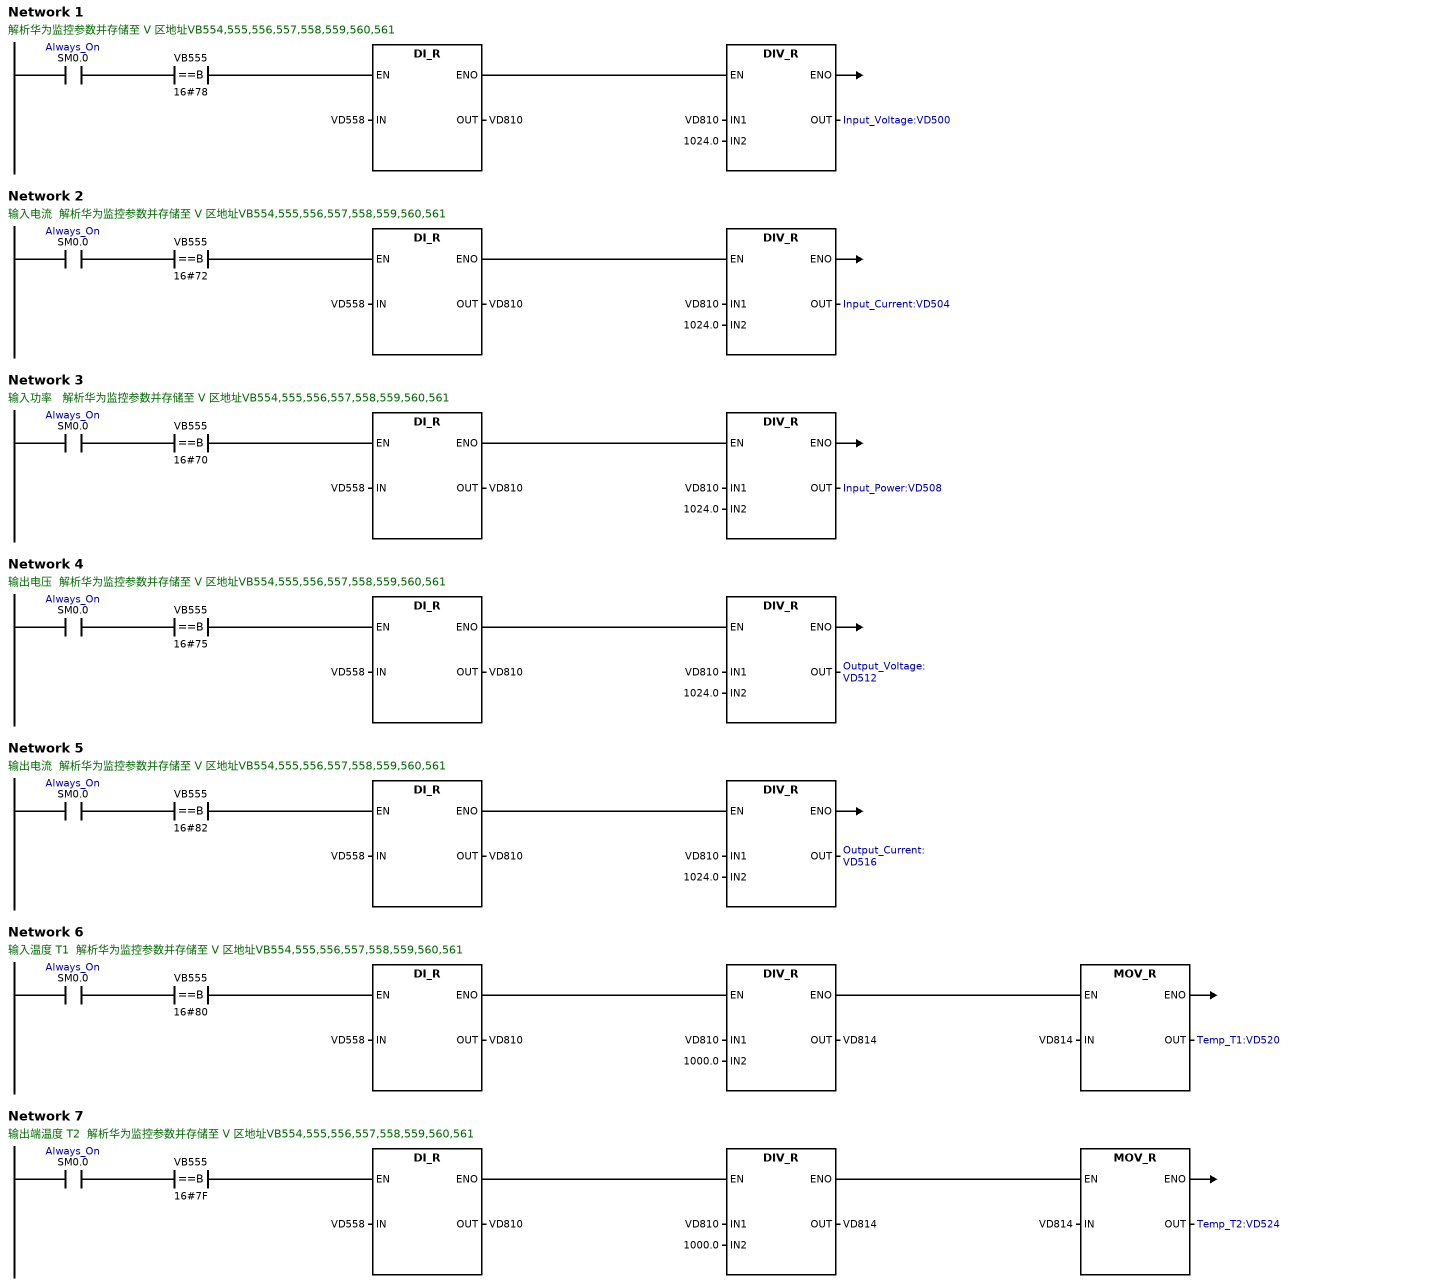
Network 1
//  解析华为监控参数并存储至 V 区地址VB554,555,556,557,558,559,560,561
// 解析标号
// 参数 ID 为 0x78 (输入电压)
// 存入 VD500 (输入电压)
LD     Always_On:SM0.0
AB=    VB555, 16#78
DTR    VD558, VD810
AENO
MOVR   VD810, Input_Voltage:VD500
/R     1024.0, Input_Voltage:VD500
Network 2
// 输入电流  解析华为监控参数并存储至 V 区地址VB554,555,556,557,558,559,560,561
// 参数 ID 为 0x72 (输入电流)
// 转换
// 缩放
// 存入 VD504 (输入电流)
LD     Always_On:SM0.0
AB=    VB555, 16#72
DTR    VD558, VD810
AENO
MOVR   VD810, Input_Current:VD504
/R     1024.0, Input_Current:VD504
Network 3
// 输入功率   解析华为监控参数并存储至 V 区地址VB554,555,556,557,558,559,560,561
// 参数 ID 为 0x70 (输入功率)
// 转换
// 缩放
// 存入 VD508 (输入功率)
LD     Always_On:SM0.0
AB=    VB555, 16#70
DTR    VD558, VD810
AENO
MOVR   VD810, Input_Power:VD508
/R     1024.0, Input_Power:VD508
Network 4
// 输出电压  解析华为监控参数并存储至 V 区地址VB554,555,556,557,558,559,560,561
// 参数 ID 为 0x75 (输出电压)
// 取值
// 缩放
// 存入 VD512 (输出电压)
LD     Always_On:SM0.0
AB=    VB555, 16#75
DTR    VD558, VD810
AENO
MOVR   VD810, Output_Voltage:VD512
/R     1024.0, Output_Voltage:VD512
Network 5
// 输出电流  解析华为监控参数并存储至 V 区地址VB554,555,556,557,558,559,560,561
// 参数 ID 为 0x82 (输出电流)
// 转换
// 缩放
// 存入 VD516 (输出电流)
LD     Always_On:SM0.0
AB=    VB555, 16#82
DTR    VD558, VD810
AENO
MOVR   VD810, Output_Current:VD516
/R     1024.0, Output_Current:VD516
Network 6
// 输入温度 T1  解析华为监控参数并存储至 V 区地址VB554,555,556,557,558,559,560,561
// 参数 ID 为 0x80 (输入温度 T1)
// 转换
// 存入 VD520 (温度 T1)
LD     Always_On:SM0.0
AB=    VB555, 16#80
DTR    VD558, VD810
AENO
MOVR   VD810, VD814
AENO
/R     1000.0, VD814
AENO
MOVR   VD814, Temp_T1:VD520
Network 7
// 输出端温度 T2  解析华为监控参数并存储至 V 区地址VB554,555,556,557,558,559,560,561
// 参数 ID 为 0x7F (输出端温度 T2)
// 转换
// 存入 VD524 (温度 T2)
LD     Always_On:SM0.0
AB=    VB555, 16#7F
DTR    VD558, VD810
AENO
MOVR   VD810, VD814
AENO
/R     1000.0, VD814
AENO
MOVR   VD814, Temp_T2:VD524
END_SUBROUTINE_BLOCK

SUBROUTINE_BLOCK SBR_3:SBR3
TITLE=控制逻辑与 IP 修改
BEGIN
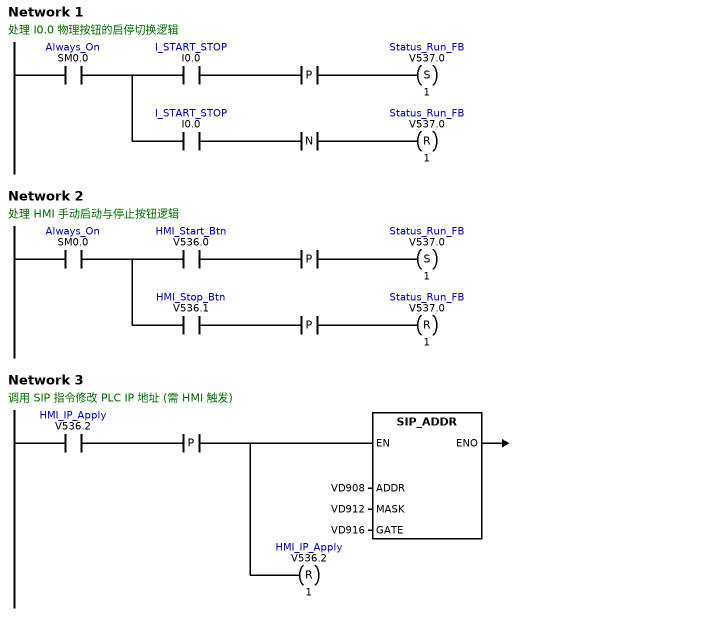
Network 1
//  处理 I0.0 物理按钮的启停切换逻辑
LD     Always_On:SM0.0
LPS
A      I_START_STOP:I0.0
EU
S      Status_Run_FB:V537.0, 1
LPP
A      I_START_STOP:I0.0
ED
R      Status_Run_FB:V537.0, 1
Network 2
//  处理 HMI 手动启动与停止按钮逻辑
LD     Always_On:SM0.0
LPS
A      HMI_Start_Btn:V536.0
EU
S      Status_Run_FB:V537.0, 1
LPP
A      HMI_Stop_Btn:V536.1
EU
R      Status_Run_FB:V537.0, 1
Network 3
//  调用 SIP 指令修改 PLC IP 地址 (需 HMI 触发)
// HMI 确认修改 IP 位
// 上升沿触发
// 应用从 VB538 开始的 IP 配置
// 位复位
LD     HMI_IP_Apply:V536.2
EU
?237   VD908, VD912, VD916
R      HMI_IP_Apply:V536.2, 1
END_SUBROUTINE_BLOCK

SUBROUTINE_BLOCK SBR_4:SBR4
TITLE=PN 通信反馈
BEGIN
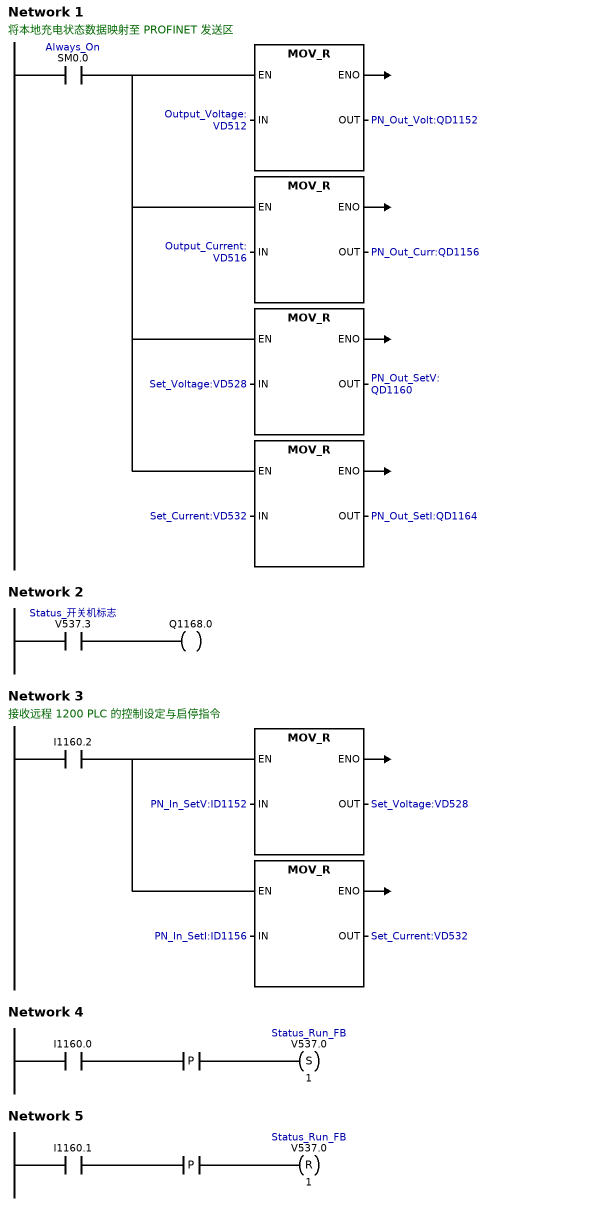
Network 1
//  将本地充电状态数据映射至 PROFINET 发送区
// 始终接通
// 实际输出电压 -> V650
// 实际输出电流 -> V654
// 当前设定电压 -> V658
// 当前设定电流 -> V662
//MOVB   VB537, PN_Out_Status        // 系统运行状态 -> V666
LD     Always_On:SM0.0
MOVR   Output_Voltage:VD512, PN_Out_Volt:QD1152
MOVR   Output_Current:VD516, PN_Out_Curr:QD1156
MOVR   Set_Voltage:VD528, PN_Out_SetV:QD1160
MOVR   Set_Current:VD532, PN_Out_SetI:QD1164
Network 2
LD     Status_开关机标志:V537.3
=      Q1168.0
Network 3
//  接收远程 1200 PLC 的控制设定与启停指令
// 始终接通
// 远程设定电压来自 V660
// 远程设定电流来自 V664
LD     I1160.2
MOVR   PN_In_SetV:ID1152, Set_Voltage:VD528
MOVR   PN_In_SetI:ID1156, Set_Current:VD532
Network 4
// 远程启动指令 (1)
// 执行启动
LD     I1160.0
EU
S      Status_Run_FB:V537.0, 1
Network 5
// 远程停止指令 (2)
// 执行停止
LD     I1160.1
EU
R      Status_Run_FB:V537.0, 1
END_SUBROUTINE_BLOCK

SUBROUTINE_BLOCK SBR_5:SBR5
TITLE=接收故障信息
BEGIN
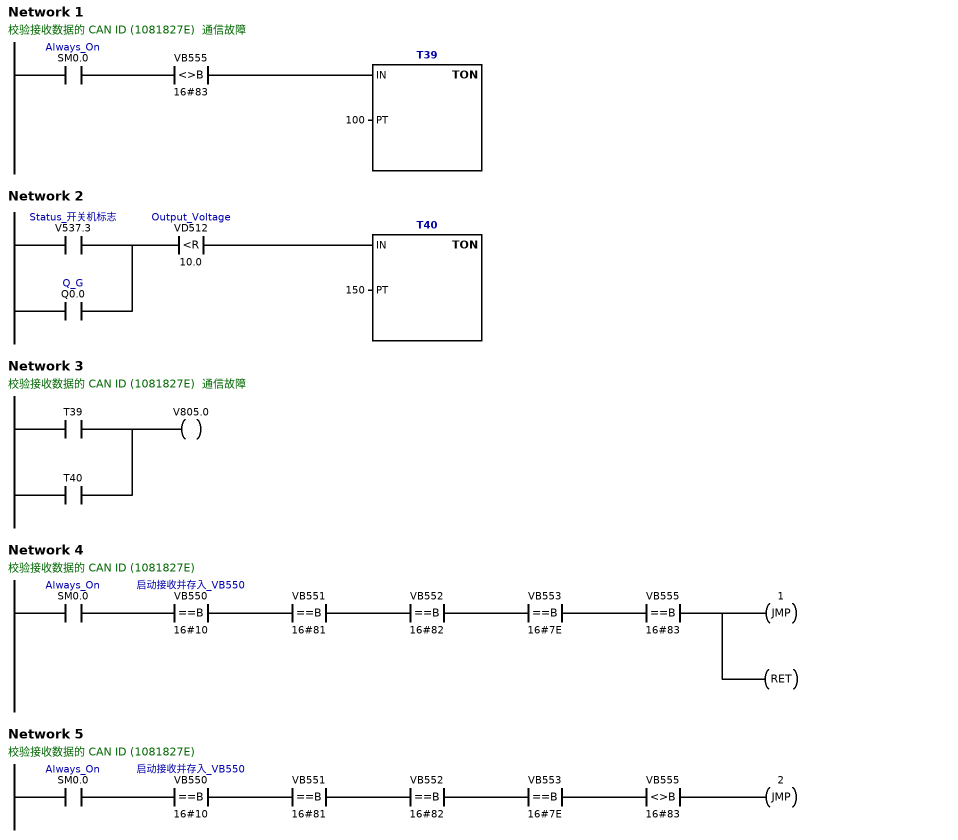
Network 1
//  校验接收数据的 CAN ID (1081827E)  通信故障
// 始终接通
// 检查 ID 字节 3
// 检查 ID 字节 2
// 检查 ID 字节 1
// 检查 ID 字节 0
// 参数 ID 为 0x83 (故障查询)
// 若匹配则跳转至解析段
LD     Always_On:SM0.0
AB<>   VB555, 16#83
TON    T39, 100
Network 2
LD     Status_开关机标志:V537.3
O      Q_G:Q0.0
AR<    Output_Voltage:VD512, 10.0
TON    T40, 150
Network 3
//  校验接收数据的 CAN ID (1081827E)  通信故障
// 始终接通
// 检查 ID 字节 3
// 检查 ID 字节 2
// 检查 ID 字节 1
// 检查 ID 字节 0
// 参数 ID 为 0x83 (故障查询)
// 若匹配则跳转至解析段
LD     T39
O      T40
=      V805.0
Network 4
//  校验接收数据的 CAN ID (1081827E)
// 始终接通
// 检查 ID 字节 3
// 检查 ID 字节 2
// 检查 ID 字节 1
// 检查 ID 字节 0
// 参数 ID 为 0x83 (故障查询)
// 若匹配则跳转至解析段
// 不匹配则退出子程序
LD     Always_On:SM0.0
AB=    启动接收并存入_VB550:VB550, 16#10
AB=    VB551, 16#81
AB=    VB552, 16#82
AB=    VB553, 16#7E
AB=    VB555, 16#83
JMP    1
CRET
Network 5
//  校验接收数据的 CAN ID (1081827E)
// 始终接通
// 检查 ID 字节 3
// 检查 ID 字节 2
// 检查 ID 字节 1
// 检查 ID 字节 0
// 参数 ID 为 0x83 (故障查询)
// 若匹配则跳转至解析段
LD     Always_On:SM0.0
AB=    启动接收并存入_VB550:VB550, 16#10
AB=    VB551, 16#81
AB=    VB552, 16#82
AB=    VB553, 16#7E
AB<>   VB555, 16#83
JMP    2
Network 6
//  解析华为故障参数并存储至 V 区地址VB554,555,556,557,558,559,560,561
LBL    1                     // 解析标号
LD     Always_On:SM0.0
MOVD   VD558, VD800          // 取出反馈数据字
Network 7
LBL    2                     // 解析标号
CRET
END_SUBROUTINE_BLOCK

// SBR6: protected block, not included

// SBR7: protected block, not included

// SBR8: protected block, not included
